TYPE ST_PortalJob :
STRUCT
	nJobID:			UDINT; //Job Nummer
	eJobType:		E_JobType;  //Neuer Stein von Stapel oder Stein auf Brett oder Stein entfernen
	fStartPosX:		LREAL; //Startposition x in mm
	fStartPosY:		LREAL; //Startposition y in mm
	fDestPosX:		LREAL; //Zielposition x in mm
	fDestPosY:		LREAL; //Zielposition y in mm
	bBlack:			BOOL; //entscheidet über Lagerposition
END_STRUCT
END_TYPE

(* stored: Version 1.1.0.1, ProductVersion 3.1.4024.12
   DUT ST_PortalJob: Id {7f9ba2e2-67a3-415e-820d-9df30c273aab} *)
